Fanuc KAREL source: ka00120.KL

-- PROVISIONAL review KL for V1013-1; original PC SHA256 796a2ed208c2bf0daa06e71c6fab5ddfb143dd598a140466ede897e8c89de4f2
-- Incomplete behavior may be omitted. Consult companion uncertainty JSON. Do not deploy.
PROGRAM KA00120
%NOLOCKGROUP
-- UNRESOLVED_DECL SRC type=00001c
-- UNRESOLVED_DECL DST type=002017
BEGIN
  -- UNRESOLVED_PC offsets 5-15; opcodes 9D,22,A5
  -- UNRESOLVED_PC offsets 20-35; opcodes 21,22,9D,33,B4
  -- UNRESOLVED_PC offsets 40-44; opcodes 7F
END KA00120
